FUNCTION_BLOCK "LModbusAscii_Master"   // FB4, SCL
TITLE = LModbusAscii_Master
{ S7_Optimized_Access := 'TRUE' }
AUTHOR : Siemens
FAMILY : LModbus
NAME : LModbusAscii_Master
VERSION : 1.1
// Modbus ASCII Master block
// the block implements the Modbus Ascii Master functionality
// ENO is not used, error handling done with error and status
   VAR_INPUT
      enable : Bool;   // True: Enables block functionality, rising edge initializes the port
      execute : Bool;   // Rising edge starts action once
      hardwareId : Hw_Any;   // Hardware Identifier for used communication module
      slaveAddress : USInt;   // Address of modbus ASCII Slave
      functionCode : USInt;   // Function code to send to the Slave
      startAddress : UInt;   // Startaddress in Modbus slave to read or write / if MB function 08, then startAddress is subfunctioncode / if MB function 43, then startAddress is object ID
      quantity : UInt;   // Quantity of Coils/Registers to read or write to /from slave device
      parameter : "LModbusAscii_typeAsciiConfiguration";   // Parameter dataset to configure modbus interface
      mask : Struct   // Logical Mask for Function Code 22 Mask Write Register
         andMask : Word;   // AND Mask of Function Code 22
         orMask : Word;   // OR Mask of Function Code 22
      END_STRUCT;
      readWrite : Struct   // Addresses and Quantities for Function Code 23 Read/Write Multiple registers
         startAddressRead : UInt := 1;   // Address to Holding Register for Read access
         quantityRead : USInt;   // Quantity of Holding Register for Read access
         startAddressWrite : UInt := 1;   // Address to Holding Register for Write access
         quantityWrite : USInt;   // Quantity of Holding Register for Write access
      END_STRUCT;
   END_VAR
   VAR_OUTPUT
      valid : Bool;   // TRUE: Valid set of output values available at the FB
      done : Bool;   // TRUE: Commanded functionality has been completed successfully
      busy : Bool;   // TRUE: FB is not finished and new output values can be expected
      error : Bool;   // TRUE: An error occurred during the execution of the FB
      status : Word := 16#7000;   // 16#0000 - 16#7FFF: Status of the FB, 16#8000 - 16#FFFF: Error identification
      diagnostics : "LModbusAscii_typeDiagnostics";   // Diagnostics information (status, subFunctionStatus, statenumber of Error)
   END_VAR
   VAR_IN_OUT
      data : Variant;   // Data for Modbus Read or Write of type Byte, Char, USInt, SInt, Bool, Word, UInt, Real, Int
   END_VAR
   VAR
      statExecuteOld : Bool;   // Old value of 'execute' input for edge detection
      statValid : Bool;   // Static value for output 'valid'
      statDone : Bool;   // Static value for output 'done'
      statBusy : Bool;   // Static value for output 'busy'
      statError : Bool;   // Static value for output 'error'
      statSerialLineStopBits : UInt;   // Serial line stop bits - defined by the parity
      statRetryCounter : USInt;   // Retry counter tag
      statFBState : DInt := 0;   // State in the state machine of the FB
      statDiagnostics : "LModbusAscii_typeDiagnostics";   // Static Diagnostic data and Information
      statEmptyDiagnostics : "LModbusAscii_typeDiagnostics";   // Empty diagnostics information (for initialization purposes only)
      statParameter : "LModbusAscii_typeAsciiConfiguration";
      instPortConfig : Port_Config;   // Instance Port configuration for Modbus ASCII Communication
      instTransmitterConfig : Send_Config;   // Instance Transmitter configuration for Modbus ASCII Communication
      instReceiverConfig : Receive_Config;   // Instance Receiver configuration for Modbus ASCII Communication
      statReceiverConditions : Receive_Conditions;   // Static Receive conditions for Modbus ASCII Communication
      instSendRequest : Send_P2P;   // Instance Send Data to Modbus slave
      instGetResponse : Receive_P2P;   // Instance Recive data from Modbus slave
      instResetRxBuffer : Receive_Reset;   // Instance Reset and clear receive buffer
      instWatchdog : IEC_TIMER;   // Instance Watchdog to check transmit to recive transition OR TurnAround delay time
      statTransmitterBuffer : Array[0..#BUFFER_UPPER_BOUND_BINARY] of Byte;   // Static Buffer for transmit data to slave device
      statReceiverBuffer : Array[0..#BUFFER_UPPER_BOUND_BINARY] of Byte;   // Static Buffer for receiving data from slave device
      statTransmitterAsciiBuffer : Array[0..#BUFFER_UPPER_BOUND_ASCII] of Byte;   // Static Buffer for the ASCII transfer string - send an receive direction
      statReceiverAsciiBuffer : Array[0..#BUFFER_UPPER_BOUND_ASCII] of Byte;   // Static Buffer for the ASCII transfer string - send an receive direction
      instAsciiDecode : "LModbusAscii_DecodeAsciiToByte";   // Instance to convert/decode the two ASCII nibble character array into byte array
      instAsciiEncode : "LModbusAscii_EncodeByteToAscii";   // Instance to convert/encode the byte array into a two ASCII nibble character array
      statReadWrite : Struct   // Addresses and Quantities for Function Code 23 Read/Write Multiple registers
         startAddressRead : UInt;
         quantityRead : USInt;
         startAddressWrite : UInt;
         quantityWrite : USInt;
      END_STRUCT;
      statHardwareId : UInt;   // Hardware Identifier for used communication module
      statErrorUserCleared : Bool;   // Error occurred that can only be solved by user; rising edge at enable input necessary
      statDisablingCompleted : Bool;   // TRUE: Disabling has been completed
      statErrorAutoCleared : Bool;   // Error occurred that can be acknowledged by FB
      statEnableOld : Bool;   // Old value of 'enable' input for edge detection
      statQuantityInBytes : USInt;   // Static internal value for quantity check in bytes
      statQuantityInBytesRead : USInt;   // Static internal value for quantity check in bytes for FC 23 Read requests
      statQuantityInBytesWrite : USInt;   // Static internal value for quantity check in bytes for FC 23 Write requests
      statFunctionCode : USInt;   // Function code to send to the Slave
      statSlaveAddress : USInt;   // Address of modbus ASCII Slave
      statQuantity : UInt;   // Static tag for quantity of requested data
      statStartAddress : UInt;   // Static tag for start address as word
      statAndMask : Word;   // AND Mask of Function Code 22
      statOrMask : Word;   // OR Mask of Function Code 22
      statLengthAfterEncoding : DInt;   // Temporary value for length of ASCII characters to transfer
      statLengthAfterDecoding : DInt;   // Temporary value for length of Byte Array received
   END_VAR
   VAR_TEMP
      tempExecute : Bool;   // Temporary value for input 'execute'
      tempStayInStatemachine : Bool;   // Temporary bool tag to stay in state machine and repeat execution if set to TRUE
      tempEnable : Bool;   // Temporary value for input 'enable'
      tempRetVal : Int;   // Temporary value for retVal of MOVE_BLK_VARIANT or DESERIALIZE
      tempSerializePos : DInt;   // Temporary value for serialize position
      tempDeserializePos : DInt;   // Temporary value for deserialize position
      tempReceiveBufferIndex : Int;   // Temporary value for receive buffer index
      tempLengthIndex : DInt;   // Temporary value for indexing buffer arrays
      tempEmptyData : Array[0..#BUFFER_UPPER_BOUND_BINARY] of Byte;   // Temporary value for reset data after disabling
      tempStartAddress : Word;   // Temporary value for Startaddress in Modbus slave to read or write / if MB function 08, then startAddress is subfunctioncode / if MB function 43, then startAddress is object ID
      tempQuantity : Word;   // Temporary value for Quantity of Coils/Registers to read or write to /from slave device
   END_VAR
   VAR CONSTANT
      FB_STATE_NO_PROCESSING_IDLE : DInt := 0;   // FB state: No processing
      FB_STATE_INIT_INTERFACE : DInt := 1;   // FB state: initialization of Port
      FB_STATE_INIT_TRANSMITTER : DInt := 2;   // FB state: initialization of Transmitter
      FB_STATE_INIT_RECEIVER : DInt := 3;   // FB state: initialization of Receiver
      FB_STATE_WAIT_FOR_EXECUTE : DInt := 4;   // FB state: wait until function should be executed
      FB_STATE_RESET_RECEIVER_BUFFER : DInt := 5;   // FB state: initialization of Receiver Buffer by clearing it
      FB_STATE_SETUP_TRANSMIT_PROTOCOL : DInt := 30;   // FB state: setup transmit protocol
      FB_STATE_TRANSMIT_DATA : DInt := 40;   // FB state: send message to slave
      FB_STATE_WAIT_FOR_RESPONSE : DInt := 41;   // FB state: wait for response from slave
      FB_STATE_WAIT_FOR_TURNAROUND_DELAY : DInt := 42;   // FB state: wait for turnaround delay after send broadcast
      FB_STATE_PROCESS_RECEIVED_DATA : DInt := 50;   // FB state: read / decode received data
      FB_STATE_DISABLING : DInt := 99;   // FB state: disabling / clear of the interface configuration
      STATUS_DONE : Word := 16#0000;   // Execution finished without errors
      STATUS_NO_CALL : Word := 16#7000;   // No job being currently processed
      STATUS_FIRST_CALL : Word := 16#7001;   // First call after enabling the block (rising edge 'enable')
      STATUS_SUBSEQUENT_CALL : Word := 16#7002;   // Subsequent call during active interface preparation without further details
      STATUS_READY : Word := 16#7003;   // Block is in ready state and waiting for a modbus job
      STATUS_EXECUTED_FIRST_CALL : Word := 16#7004;   // First call after incoming new job (rising edge 'execute')
      STATUS_EXECUTED_SUBSEQUENT_CALL : Word := 16#7005;   // Subsequent call during active job processing without further details
      NO_ERROR : Word := 16#0000;   // Blank error code / no error
      ERR_UNDEFINED_STATE : Word := 16#8600;   // Error due to an undefined state in state machine
      ERR_MODBUS_ADDRESS_OUT_OF_RANGE : Word := 16#8601;   // Error due to missconfiguration, Modbus address out of range 0 <= Address <= 247
      ERR_MODBUS_WRONG_PARITY_MODE : Word := 16#8602;   // Error due to missconfiguration, Modbus parity mode can be even(2), odd(3), no parity(1)
      ERR_MODBUS_WRONG_INTERFACE_MODE : Word := 16#8603;   // Error due to missconfiguration, Serial interface mode can be serial interface mode 0/FullDuplex (RS232), 4/Half duplex (RS485, two-wire mode)
      ERR_CONFIGURATION_PORT : Word := 16#8604;   // Error due to Port configuration, please check subfunction status in Diagnostic
      ERR_CONFIGURATION_TRANSMITTER : Word := 16#8605;   // Error due to Transmitter configuration, please check subfunction status in Diagnostic
      ERR_CONFIGURATION_RECEIVER : Word := 16#8606;   // Error due to Receiver configuration, please check subfunction status in Diagnostic
      ERR_CLEAR_RECEIVER_BUFFER : Word := 16#8607;   // Error due to clear Receiver buffer, please check subfunction status in Diagnostic
      ERR_MOVE_BLK_VAR_TO_DATA : Word := 16#8608;   // Error due to moving received data to INOUT data
      ERR_DESERIALIZE_TO_DATA : Word := 16#8609;   // Error due to deserializing received data to INOUT data
      ERR_REQUEST_NOT_SUPPORTED_FUNCTION_CODE : Word := 16#8610;   // Error due to given Modbus Function Code, not supported function, see subFctStatus in diagnostic
      ERR_REQUEST_INVALID_FC08_REQUEST_DATA : Word := 16#8681;   // Error due to given request data - for function code 8 / sub function code 1 data field needs to be 16#0000 (leave log) or 16#FF00 (clear log)
      ERR_RESPONSE_NOT_SUPPORTED_FUNCTION_CODE : Word := 16#8620;   // Error due to received Modbus Function Code, not supported function, see subFctStatus in diagnostic
      ERR_INTERFACE_NOT_CONFIGURED : Word := 16#8611;   // Error due to interface, that was not configured yet
      ERR_SERIALIZE_MULTIPLE_WRITE : Word := 16#8612;   // Error due to serializing data to transmitter buffer at multiple write request
      ERR_SERIALIZE_SINGLE_WRITE : Word := 16#8622;   // Error due to serializing data to transmitter buffer at single write request
      ERR_MOVE_BLK_VAR_MULTIPLE_WRITE : Word := 16#8613;   // Error due to moving data to transmitter buffer
      ERR_INVALID_QUANTITY : Word := 16#8615;   // Error due to invalid quantity for read (125) or write (121) request
      ERR_MOVE_BLK_VAR_RECEIVE_DATA : Word := 16#8633;   // Error due to moving receive buffer to data
      ERR_MOVE_BLK_VAR_SINGLE_WRITE : Word := 16#8623;   // Error due to moving data to transmitter buffer
      ERR_DATA_TYPE_NOT_SUPPORTED : Word := 16#8614;   // Error due to moving data to INOUT data. Has to be Array of Byte or Word.
      ERR_TRANSMISSION_FAILURE : Word := 16#8201;   // Error during data transmisson to slave, please check subfunction status in Diagnostic
      ERR_RESPONSE_TIMEOUT_EXPIRATION : Word := 16#8202;   // Error due to timeout while wait for response from slave, "response time-out expiration"
      ERR_RECEIVER_FAILURE : Word := 16#8203;   // Error due to receiver data from slave, please check subfunction status in Diagnostic
      ERR_RESPONSE_EXCEPTION_FROM_SLAVE : Word := 16#8204;   // Error due to an received exception from slave - excpetion code is stored in diagnostics subFunctionStatus
      ERR_RESPONSE_WRONG_LRC : Word := 16#8205;   // Error due to LRC Check on response data
      ERR_RESPONSE_WRONG_QUANTITY : Word := 16#8206;   // Error due to wrong quantity received
      ERR_RESPONSE_SINGLE_WRITE : Word := 16#8207;   // Error due to response of single write functions
      ERR_RESPONSE_MULTI_WRITE : Word := 16#8217;   // Error due to response of multiple write functions
      ERR_RESPONSE_NOT_EXPECTED_FC : Word := 16#8208;   // Error because response contains not expected function code
      ERR_RESPONSE_NOT_EXPECTED_SUB_FC : Word := 16#8218;   // Error because response contains not expected subfunction code
      ERR_RESPONSE_WRONG_SLAVE : Word := 16#8209;   // Error due to wrong slave answered to request
      ERR_NOT_SUPPORTED_SUB_FC : Word := 16#8210;   // Error due to not supported function code for diagnostic function 08
      ERR_DIAG_SUB_0 : Word := 16#8250;   // Error in response for diagnostic subfunction 0 (Return query value) - wrong echo value
      ERR_DIAG_SUB_1 : Word := 16#8251;   // Error in response for diagnostic subfunction 1 (Restart Com) - wrong echo value
      FREEPORT_PROTOCOL : UInt := 0;   // Freeport protocol is used for Modbus ASCII
      FB_DISABLE_TIME : Time := T#500Ms;   // Time that any active instances may need until the device is hard deactivated.
      BUFFER_UPPER_BOUND_ASCII : DInt := 608;   // Upper Bound of Buffer ASCII Char mode
      BUFFER_UPPER_BOUND_BINARY : DInt := 300;   // Upper Bound of Buffer in Byte to store the binary data
      DATA_INDEX_0 : Int := 0;   // Data index set to 0
      INITIALIZE_WORD_0 : Word := 16#0000;   // Initialize Word (16#00)
      B1_OFFSET : USInt := 1;   // Offset to select high byte in a word
      FC05_SET_COMMAND_IDENT : Word := 16#FF00;   // Modbus ASCII - identifier for setting coil to true
      MODBUS_INTERFACE_MODE_RS232 : USInt := 0;   // Modbus interface modus is RS232 Full Duplex
      MODBUS_INTERFACE_MODE_RS485 : USInt := 4;   // Modbus interface modus is RS485 Half Duplex
      MODBUS_ADDRESS_MAX : USInt := 247;   // Modbus ASCII maximum address range is 247
      MODBUS_ADDRESS_BROADCAST : USInt := 0;   // Modbus ASCII broadcast address is 0
      MODBUS_ASCII_SEVEN_DATABITS : UInt := 2;   // Modbus ASCII Databits defined --> 7
      MODBUS_ASCII_PARITY_EVEN : UInt := 2;   // Modbus ASCII EVEN Parity setting for port configuration
      MODBUS_ASCII_PARITY_ODD : UInt := 3;   // Modbus ASCII ODD Parity setting for port configuration
      MODBUS_ASCII_NO_PARITY : UInt := 1;   // Modbus ASCII NO Parity setting for port configuration
      MODBUS_ASCII_STOPBITS_NO_PARITY : UInt := 2;   // Modbus ASCII Stopbits = 2 if no parity mode is choosen
      MODBUS_ASCII_STOPBITS_WITH_PARITY : UInt := 1;   // Modbus ASCII Stopbits = 1 if even or odd parity mode is choosen
      MODBUS_TURNAROUND_DELAY : Time := T#200MS;   // Modbus turnaround delay time after a broadcast request was send
      MODBUS_SLAVE_ADDRESS_INDEX : USInt := 0;   // Modbus Master / Slave request / response - index for slave address
      MODBUS_FUNCTION_CODE_INDEX : USInt := 1;   // Modbus Master / Slave request / response - index for function code AND Exception notice (MSB) in response buffer
      MODBUS_RESPONSE_BYTE_COUNT_INDEX : USInt := 2;   // Modbus Master - Index to length entry in response field
      MODBUS_RESPONSE_ADDRESS_INDEX : USInt := 2;   // Modbus Master - Index to start address in response field
      MODBUS_RESPONSE_QUANTITY_INDEX : USInt := 4;   // Modbus Master - Index to quantity in response field
      MODBUS_EXCEPTION_CODE_INDEX : USInt := 1;   // Modbus Slave response - index for exception code in response buffer
      MODBUS_DEFAULT_REQUEST_LENGTH : USInt := 2;   // Modbus Master request - shortest possible request length
      MODBUS_DEFAULT_RESP_INDEX : USInt := 2;   // Modbus Master response - default response index
      MODBUS_STARTADDRESS_INDEX : USInt := 2;   // Modbus Master request - index for start address
      MODBUS_STARTADDRESS_FC23_WRITE_INDEX : USInt := 6;   // Modbus Master request - index for start address of write job for FC 23 request
      MODBUS_AND_MASK_INDEX : USInt := 4;   // Modbus Master request - index for AND Mask for fc 22
      MODBUS_OR_MASK_INDEX : USInt := 6;   // Modbus Master request - index for OR Mask for fc 22
      MODBUS_QUANTITY_INDEX : USInt := 4;   // Modbus Master request - index for quantity
      MODBUS_QUANTITY_FC23_WRITE_INDEX : USInt := 8;   // Modbus Master request - index for quantity of write job for FC 23 request
      MODBUS_BYTE_COUNT_INDEX : USInt := 6;   // Modbus Master request - index byte count
      MODBUS_BYTE_COUNT_FC23_INDEX : USInt := 10;   // Modbus Master request - index byte count of write job for FC 23 request
      MODBUS_DATA_INDEX : USInt := 7;   // Modbus Master request - index to first data entry
      MODBUS_FC23_DATA_INDEX : USInt := 11;   // Modbus Master request - index to first data entry of write job for FC 23 request
      MODBUS_USER_DATA_READ_INDEX : USInt := 3;   // Modbus Slave response - index for position of user data
      MODBUS_DIAG_SUB_FC_INDEX : USInt := 2;   // Modbus Master / Slave request / Response - index for subfunction code at Diagnostic function and Device ident
      MODBUS_DIAG_DATA_INDEX : USInt := 4;   // Modbus Master / Slave request / Response - index for subfunction code at Diagnostic function and Device ident
      MODBUS_REQUEST_LENGTH : UInt := 6;   // Modbus Master request length
      MODBUS_REQUEST_MULTIPLE_WRITE_LENGTH : UInt := 7;   // Modbus Master request length for multiple write functions
      MODBUS_REQUEST_MASK_WRITE_LENGTH : UInt := 8;   // Modbus Master request length for mask write function
      MODBUS_REQUEST_READ_WRITE_LENGTH : UInt := 11;   // Modbus Master request length for FC 23 read/write request
      MODBUS_STARTADDRESS_CORRECTION : USInt := 1;   // Correction of MODBUS startaddress by subtraction of 1
      MODBUS_MAX_REGISTER_READ : USInt := 125;   // Modbus maximum quantity for register read requests
      MODBUS_MAX_REGISTER_WRITE : USInt := 123;   // Modbus maximum quantity for register write requests
      MODBUS_FC23_MAX_REGISTER_WRITE : USInt := 121;   // Modbus maximum quantity for FC 23 register write requests
      MODBUS_FC43_MEI_TYE : Byte := 16#0E;   // Modbus MEI Type for Device Identification
      MODBUS_FC43_DEVICE_ID_CODE_INDEX : USInt := 3;   // Modbus Device ID code index in request
      MODBUS_FC43_OBJECT_ID_CODE_INDEX : USInt := 4;   // Modbus Object ID code index in request
      MODBUS_FC43_REQUEST_LENGTH : USInt := 5;   // Modbus Master request length for FC 43 request
      MB_FC_01_READ_COILS : USInt := 1;   // Modbus function code 01 - read coils
      MB_FC_02_READ_DISCRETE_INPUTS : USInt := 2;   // Modbus function code 02 - read discrete inputs
      MB_FC_03_READ_HOLDING_REGISTERS : USInt := 3;   // Modbus function code 03 - read holding registers
      MB_FC_04_READ_INPUT_REGISTERS : USInt := 4;   // Modbus function code 04 - read input registers
      MB_FC_05_WRITE_COIL : USInt := 5;   // Modbus function code 05 - write single coil
      MB_FC_06_WRITE_REGISTER : USInt := 6;   // Modbus function code 06 - write single register
      MB_FC_07_READ_EXCEPTION_STATUS : USInt := 7;   // Modbus function code 07 - read exception status
      MB_FC_08_DIAGNOSTIC : USInt := 8;   // Modbus function code 08 - diagnostic
      MB_FC_11_GET_COM_EVENT_COUNTER : USInt := 11;   // Modbus function code 11 - diagnostic
      MB_FC_12_GET_COM_EVENT_LOG : USInt := 12;   // Modbus function code 12 - get comm event log
      MB_FC_15_WRITE_COILS : USInt := 15;   // Modbus function code 15 - write multiple coils
      MB_FC_16_WRITE_REGISTERS : USInt := 16;   // Modbus function code 16 - write multiple registers
      MB_FC_22_MASK_WRITE_REGISTER : USInt := 22;   // Modbus function code 22 - mask Write Register
      MB_FC_23_READ_WRITE_MULTIPLE_REGISTERS : USInt := 23;   // Modbus function code 23 - read/write Multiple registers
      MB_FC_43_READ_DEVICE_IDENT : USInt := 43;   // Modbus function code 43 - read device idendification data
      DIAG_SUB_FC_0_RETURN_QUERY_DATA : USInt := 16#00;   // Diag: Return query dara
      DIAG_SUB_FC_1_RESTART_COM : USInt := 16#01;   // Diag: Restart communication option
      DIAG_SUB_FC_2_RETURN_DIAG_REGISTER : USInt := 16#02;   // Diag: Return diagnostic register
      DIAG_SUB_FC_4_FORCE_LISTEN_ONLY : USInt := 16#04;   // Diag: Force listen only
      DIAG_SUB_FC_10_CLEAR_DIAG_REGISTER : USInt := 16#0A;   // Diag: Clear counter and diagnostic register
      DIAG_SUB_FC_11_COUNTER_TOTAL_MESSAGE : USInt := 16#0B;   // Diag: Return bus message count
      DIAG_SUB_FC_12_COUNTER_CRC_ERR : USInt := 16#0C;   // Diag: Return bus commuunication error count
      DIAG_SUB_FC_13_COUNTER_EXCEPTION_ERR : USInt := 16#0D;   // Diag: Return bus exception error count
      DIAG_SUB_FC_14_COUNTER_TOTAL_MESSAGES : USInt := 16#0E;   // Diag: Return server message count
      DIAG_SUB_FC_15_COUNTER_NO_RESPONSE : USInt := 16#0F;   // Diag: Return Server no respomse count
      DIAG_SUB_FC_16_COUNTER_NAK : USInt := 16#10;   // Diag: Return Server negative acknowledge count
      DIAG_SUB_FC_17_COUNTER_SERVER_BUSY : USInt := 16#11;   // Diag: Return Server busy count
      DIAG_SUB_FC_18_BUS_CHAR_OVERRUN : USInt := 16#12;   // Diag: Return Bus Character Overrun Count
      DIAG_SUB_FC_20_CLEAR_OVERRUN : USInt := 16#14;   // Diag: Clear Overrun Counter and Flag
   END_VAR
   // statDiagnostics.status := 16#7000;
BEGIN
   REGION BLOCK INFO HEADER
     //===============================================================================
     // SIEMENS / (c)copyright 2026
     //-------------------------------------------------------------------------------
     // Title:            LModbusAscii_Master
     // Comment/Function: Modbus ASCII Master
     //                   The block implements the Modbus ASCII Master functionality.
     //                   ENO is not used, error handling done with error and status.
     // Library/Family:   LModbus
     // Author:           Siemens
     // Tested with:      S7-1200/1500
     // Engineering:      TIA Portal >= V19
     // Restrictions:     (none)
     // Requirements:     CM (RS485)
     //-------------------------------------------------------------------------------
     // Change log table:
     // Version  | Date       | Expert in charge       | Changes applied
     //----------|------------|------------------------|------------------------------
     // 00.01.00 | 2019-08-05 | Siemens                | first released version
     // 01.00.00 | 2023-03-20 | Siemens                | Styleguide adaptions and bugfix for data output
     // 01.01.00 | 2026-05-29 | Siemens                | New Functions and BugFix
     //===============================================================================
   END_REGION

   REGION ENABLING/DISABLING
     #tempEnable := #enable; // work with temporary value
     #tempExecute := #execute; // work with temporary value

     IF (#tempEnable = TRUE) AND (#statDiagnostics.status = #STATUS_NO_CALL) THEN // Enable FB
       REGION Enable
         // first call; initialize FB
         REGION Initialize standard interface
           #statBusy := TRUE;
           #statError := FALSE;
           #statErrorUserCleared := FALSE;
           #statErrorAutoCleared := FALSE;
           #statDiagnostics.status := #STATUS_FIRST_CALL;
           #statDiagnostics.subFunctionStatus := #NO_ERROR;
           #statDiagnostics.stateNumber := 0;
           #diagnostics := #statEmptyDiagnostics;
           #statDisablingCompleted := FALSE;
         END_REGION Initialize standard interface

         REGION Verify Input parameters
           #statParameter := #parameter;
           // verify interface mode is RS232 or RS485
           IF #statParameter.modeInterfacePTP <> #MODBUS_INTERFACE_MODE_RS232
             AND #statParameter.modeInterfacePTP <> #MODBUS_INTERFACE_MODE_RS485
           THEN
             #statErrorUserCleared := TRUE;
             #statDiagnostics.status := #ERR_MODBUS_WRONG_INTERFACE_MODE;

             // check parity mode even odd or non parity
           ELSIF #statParameter.parity <> #MODBUS_ASCII_NO_PARITY
             AND #statParameter.parity <> #MODBUS_ASCII_PARITY_EVEN
             AND #statParameter.parity <> #MODBUS_ASCII_PARITY_ODD
           THEN
             #statErrorUserCleared := TRUE;
             #statDiagnostics.status := #ERR_MODBUS_WRONG_PARITY_MODE;
           END_IF;

           #statHardwareId := #hardwareId;
         END_REGION

         REGION Init static tags
           // adjust stop bits for serial interface configuration
           IF #statParameter.parity = #MODBUS_ASCII_NO_PARITY THEN
             // if no Parity is choosen, two stop bits are needed
             #statSerialLineStopBits := #MODBUS_ASCII_STOPBITS_NO_PARITY;
           ELSE
             // if even or odd Parity is choosen, just one stop bit is needed
             #statSerialLineStopBits := #MODBUS_ASCII_STOPBITS_WITH_PARITY;
           END_IF;
         END_REGION Init static tags

         REGION Init instances by call subsidiary FBs with false
           #instPortConfig(REQ := FALSE);
           #instTransmitterConfig(REQ := FALSE);
           #instReceiverConfig(REQ := FALSE,
                               Receive_Conditions := #statReceiverConditions);
           #instSendRequest(REQ := FALSE,
                            BUFFER:=#statTransmitterAsciiBuffer);
         END_REGION Init instances by call subsidiary FBs with false

         // state machine - start functionality
         #statFBState := #FB_STATE_INIT_INTERFACE;
       END_REGION Enable

     ELSIF (#tempEnable = FALSE) AND (#statEnableOld = TRUE) THEN // disable FB 
       REGION Disable
         #statFBState := #FB_STATE_DISABLING;
         #instWatchdog.TON(IN := FALSE, PT := #FB_DISABLE_TIME);
       END_REGION Disable

     ELSIF (#statDiagnostics.status = #STATUS_FIRST_CALL) THEN // set status identifier of subsequent call
       REGION Subsequent
         #statDiagnostics.status := #STATUS_SUBSEQUENT_CALL;
       END_REGION Subsequent

     ELSIF NOT #tempEnable
       AND #statDiagnostics.status = #STATUS_NO_CALL
       AND (#tempExecute = TRUE)
       AND (#statExecuteOld = FALSE) // check if FB is triggered
     THEN
       REGION Faulty Call - execute with disabled function block
         #statErrorUserCleared := TRUE;
         #statDiagnostics.status := #ERR_INTERFACE_NOT_CONFIGURED;
         #statDiagnostics.subFunctionStatus := #NO_ERROR;
       END_REGION Faulty Call - execute with disabled function block

     END_IF;

     // edge detection 'enable' input
     #statEnableOld := #tempEnable;
   END_REGION ENABLING/DISABLING

   IF (#statDiagnostics.status = #STATUS_NO_CALL) THEN // nothing to do -> End here to reduce "system load"
     RETURN;
   END_IF;

   REGION STATE_MACHINE
     REPEAT
       // set repeat condition to FALSE to leave state machine loop
       #tempStayInStatemachine := FALSE;
       CASE #statFBState OF // state machine of FB
         #FB_STATE_NO_PROCESSING_IDLE: // no processing active (Note: this state must always be present and left empty)
           REGION No Processing
             ;
           END_REGION No Processing

         #FB_STATE_INIT_INTERFACE:
           REGION Init Interface
             // call port configuration to set parameters for communication
             #instPortConfig(REQ := TRUE,
                             "PORT" := #statHardwareId,
                             PROTOCOL := #FREEPORT_PROTOCOL,
                             BAUD := #statParameter.baud,
                             PARITY := #statParameter.parity,
                             DATABITS := #MODBUS_ASCII_SEVEN_DATABITS,
                             STOPBITS := #statSerialLineStopBits,
                             MODE := #statParameter.modeInterfacePTP);

             // port configuration finished successfully
             IF (#instPortConfig.DONE = TRUE) THEN
               #instPortConfig(REQ := FALSE);  // reset port config REQ input after call
               #statFBState := #FB_STATE_INIT_TRANSMITTER;   // set next state

               // error occurred during Port Configuration
             ELSIF (#instPortConfig.ERROR = TRUE) THEN
               // write diagnostic Information
               #statErrorUserCleared := TRUE;
               #statDiagnostics.status := #ERR_CONFIGURATION_PORT; // set correct status that identifies error clearly
               #statDiagnostics.subFunctionStatus := #instPortConfig.STATUS; // status of Port Configuration
               #statDiagnostics.stateNumber := #statFBState; // set error state number for diagnostic

               #instPortConfig(REQ := FALSE); // reset port config REQ input after call
             END_IF;
           END_REGION Init Interface

         #FB_STATE_INIT_TRANSMITTER:
           REGION Init Transmitter
             // call transmitter configuration to set paramters for communication (SEND_CFG)
             #instTransmitterConfig(REQ := TRUE,
                                    "PORT" := #statHardwareId);

             // port configuration finished successfully
             IF (#instTransmitterConfig.DONE = TRUE) THEN
               #instTransmitterConfig(REQ := FALSE);   // reset receiver config REQ input after call
               #statFBState := #FB_STATE_INIT_RECEIVER;  // set next state

               // error occurred during Port Configuration
             ELSIF (#instTransmitterConfig.ERROR = TRUE) THEN
               // write diagnostic Information
               #statErrorUserCleared := TRUE;
               #statDiagnostics.status := #ERR_CONFIGURATION_TRANSMITTER; // set correct status that identifies error clearly
               #statDiagnostics.subFunctionStatus := #instTransmitterConfig.STATUS; // status of Port Configuration
               #statDiagnostics.stateNumber := #statFBState; // set error state number for diagnostic

               #instTransmitterConfig(REQ := FALSE); // reset receiver config REQ input after call
             END_IF;
           END_REGION Init Transmitter

         #FB_STATE_INIT_RECEIVER:
           REGION Init Receiver
             // call receiver configuration to set paramters for communication (RCV_CFG)
             #instReceiverConfig(REQ := TRUE,
                                 "PORT" := #statHardwareId,
                                 Receive_Conditions := #statReceiverConditions);

             // port configuration finished successfully
             IF (#instReceiverConfig.DONE = TRUE) THEN
               #instReceiverConfig(REQ := FALSE,
                                   Receive_Conditions := #statReceiverConditions); // reset receiver config REQ input after call

               #statValid := TRUE;
               #statBusy := FALSE;
               #statDiagnostics.status := #STATUS_READY;
               #statFBState := #FB_STATE_WAIT_FOR_EXECUTE; // set next state

               // error occurred during Port Configuration
             ELSIF (#instReceiverConfig.ERROR = TRUE) THEN
               // write diagnostic Information
               #statErrorUserCleared := TRUE;
               #statDiagnostics.status := #ERR_CONFIGURATION_RECEIVER; // set correct status that identifies error clearly
               #statDiagnostics.subFunctionStatus := #instReceiverConfig.STATUS; // status of Port Configuration
               #statDiagnostics.stateNumber := #statFBState; // set error state number for diagnostic

               #instReceiverConfig(REQ := FALSE,
                                   Receive_Conditions := #statReceiverConditions); // reset receiver config REQ input after call
             END_IF;
           END_REGION Init Receiver

         #FB_STATE_WAIT_FOR_EXECUTE:
           REGION Wait for execute
             REGION Execute
               IF (#tempExecute = TRUE) AND (#statExecuteOld = FALSE) // check if FB is triggered
               THEN
                 REGION Verify input paramters
                   #statFunctionCode := #functionCode;
                   #statSlaveAddress := #slaveAddress;

                   // check, if requested function code is supported by the function block
                   IF #statFunctionCode <> #MB_FC_01_READ_COILS
                     AND #statFunctionCode <> #MB_FC_02_READ_DISCRETE_INPUTS
                     AND #statFunctionCode <> #MB_FC_03_READ_HOLDING_REGISTERS
                     AND #statFunctionCode <> #MB_FC_04_READ_INPUT_REGISTERS
                     AND #statFunctionCode <> #MB_FC_05_WRITE_COIL
                     AND #statFunctionCode <> #MB_FC_06_WRITE_REGISTER
                     AND #statFunctionCode <> #MB_FC_07_READ_EXCEPTION_STATUS
                     AND #statFunctionCode <> #MB_FC_08_DIAGNOSTIC
                     AND #statFunctionCode <> #MB_FC_11_GET_COM_EVENT_COUNTER
                     AND #statFunctionCode <> #MB_FC_12_GET_COM_EVENT_LOG
                     AND #statFunctionCode <> #MB_FC_15_WRITE_COILS
                     AND #statFunctionCode <> #MB_FC_16_WRITE_REGISTERS
                     AND #statFunctionCode <> #MB_FC_22_MASK_WRITE_REGISTER
                     AND #statFunctionCode <> #MB_FC_23_READ_WRITE_MULTIPLE_REGISTERS
                     AND #statFunctionCode <> #MB_FC_43_READ_DEVICE_IDENT
                   THEN
                     REGION invalid function code
                       // FB stays in wait for execute state and can be triggerde again with supported function code
                       #statErrorAutoCleared := TRUE;
                       #statDiagnostics.status := #ERR_REQUEST_NOT_SUPPORTED_FUNCTION_CODE;
                       #statDiagnostics.subFunctionStatus := USINT_TO_WORD(#statFunctionCode); // Given function code
                       #statDiagnostics.stateNumber := #statFBState; // Set error state number for diagnostic
                       EXIT; //end of block
                     END_REGION invalid function code

                   ELSIF #statSlaveAddress > #MODBUS_ADDRESS_MAX THEN
                     REGION invalid slave address
                       // verify Modbus address exceeds maximum address range
                       #statErrorAutoCleared := TRUE;
                       #statDiagnostics.subFunctionStatus := USINT_TO_WORD(#statSlaveAddress);
                       #statDiagnostics.status := #ERR_MODBUS_ADDRESS_OUT_OF_RANGE;
                       #statDiagnostics.stateNumber := #statFBState;
                       EXIT;
                     END_REGION invalid slave address

                   ELSE
                     REGION initialize function code
                       // set internal retry counter
                       // copy number of retries for retry transmition counter
                       #statRetryCounter := #statParameter.numberOfRetries;

                       // initialize statQuantity and statStartAddress
                       #statQuantity := #quantity;
                       #statStartAddress := #startAddress;

                       // check requested quantity. Later this value will be compared with the received data
                       IF #statFunctionCode = #MB_FC_01_READ_COILS
                         OR #statFunctionCode = #MB_FC_02_READ_DISCRETE_INPUTS
                         OR #statFunctionCode = #MB_FC_15_WRITE_COILS
                       THEN
                         //parameter quantity means count of bits. Eight bits are one bytes long
                         #statQuantityInBytes := UINT_TO_USINT(#statQuantity / 8);
                         IF #statQuantity MOD 8 <> 0 THEN
                           #statQuantityInBytes += 1;
                         END_IF;

                       ELSIF #statFunctionCode = #MB_FC_03_READ_HOLDING_REGISTERS
                         OR #statFunctionCode = #MB_FC_04_READ_INPUT_REGISTERS
                         OR #statFunctionCode = #MB_FC_16_WRITE_REGISTERS
                       THEN
                         // parameter quantity means count of registers. One register is two bytes long
                         #statQuantityInBytes := UINT_TO_USINT(#statQuantity) * 2;

                       ELSIF (#statFunctionCode = #MB_FC_08_DIAGNOSTIC AND #statQuantity <> #DIAG_SUB_FC_4_FORCE_LISTEN_ONLY)
                         OR #statFunctionCode = #MB_FC_05_WRITE_COIL
                         OR #statFunctionCode = #MB_FC_06_WRITE_REGISTER
                         OR #statFunctionCode = #MB_FC_07_READ_EXCEPTION_STATUS
                       THEN
                         // two bytes fixed for reply request (ping behaviour) and for single register and coil write 
                         #statQuantityInBytes := 2;

                       ELSIF #statFunctionCode = #MB_FC_22_MASK_WRITE_REGISTER THEN
                         #statQuantityInBytes := 0;
                         #statAndMask := #mask.andMask;
                         #statOrMask := #mask.orMask;

                       ELSIF #statFunctionCode = #MB_FC_23_READ_WRITE_MULTIPLE_REGISTERS THEN
                         #statReadWrite.startAddressRead := #readWrite.startAddressRead;
                         #statReadWrite.quantityRead := #readWrite.quantityRead;
                         #statReadWrite.startAddressWrite := #readWrite.startAddressWrite;
                         #statReadWrite.quantityWrite := #readWrite.quantityWrite;
                         #statQuantityInBytesRead := #statReadWrite.quantityRead * 2;
                         #statQuantityInBytesWrite := #statReadWrite.quantityWrite * 2;

                       ELSIF #statFunctionCode = #MB_FC_11_GET_COM_EVENT_COUNTER THEN
                         #statQuantityInBytes := 4;

                       ELSIF #statFunctionCode = #MB_FC_43_READ_DEVICE_IDENT THEN
                         #statQuantityInBytes := 250;
                       END_IF;
                     END_REGION initialize function code

                   END_IF;

                 END_REGION Verify input paramters

                 REGION Init instances by call subsidiary FBs with FALSE
                   #instResetRxBuffer(REQ := FALSE,
                                      "PORT" := #statHardwareId);
                   #instWatchdog.TON(IN := FALSE,
                                     PT := #statParameter.transmissionWatchdog);
                 END_REGION Init instances by call subsidiary FBs with FALSE

                 // state machine - start processing
                 #statBusy := TRUE;
                 #statFBState := #FB_STATE_RESET_RECEIVER_BUFFER;
                 #statDiagnostics.status := #STATUS_EXECUTED_FIRST_CALL;

               ELSIF NOT #tempExecute AND #statDone THEN
                 #statDiagnostics.status := #STATUS_READY;
                 #statDone := FALSE;
                 #statError := FALSE;
               END_IF;

               // edge detection 'execute' input
               #statExecuteOld := #tempExecute;
             END_REGION Execute
           END_REGION

         #FB_STATE_RESET_RECEIVER_BUFFER:
           REGION Reset Receiver Buffer
             IF #statDiagnostics.status = #STATUS_EXECUTED_FIRST_CALL THEN
               #statDiagnostics.status := #STATUS_EXECUTED_SUBSEQUENT_CALL;
             END_IF;

             // call receiver reset buffer to clear it
             #instResetRxBuffer(REQ := TRUE,
                                "PORT" := #statHardwareId);

             // port configuration finished successfully
             IF (#instResetRxBuffer.DONE = TRUE) THEN
               #instResetRxBuffer(REQ := FALSE);   // reset receiver config REQ input after call
               #statFBState := #FB_STATE_SETUP_TRANSMIT_PROTOCOL;  // set next state

               // error occurred during Port Configuration
             ELSIF (#instResetRxBuffer.ERROR = TRUE) THEN
               // write diagnostic Information
               #statErrorAutoCleared := TRUE;
               #statDiagnostics.status := #ERR_CLEAR_RECEIVER_BUFFER; // set correct status that identifies error clearly
               #statDiagnostics.subFunctionStatus := #instResetRxBuffer.STATUS; // status of Port Configuration
               #statDiagnostics.stateNumber := #statFBState; // set error state number for diagnostic

               #instResetRxBuffer(REQ := FALSE);   // reset receiver config REQ input after call
             END_IF;
           END_REGION Init Receiver Buffer

         #FB_STATE_SETUP_TRANSMIT_PROTOCOL:
           REGION Setup Transmit Protocol
             // set up communication Buffer
             // first part: is the address
             #statTransmitterBuffer[#MODBUS_SLAVE_ADDRESS_INDEX] := USINT_TO_BYTE(#statSlaveAddress);
             // second part: is the function code
             #statTransmitterBuffer[#MODBUS_FUNCTION_CODE_INDEX] := USINT_TO_BYTE(#statFunctionCode);
             // third part: set start address for request

             IF #statFunctionCode <> #MB_FC_08_DIAGNOSTIC AND #statFunctionCode <> #MB_FC_43_READ_DEVICE_IDENT THEN
               #statStartAddress := #statStartAddress - #MODBUS_STARTADDRESS_CORRECTION;
             END_IF;

             // third part: tx / transmit data protocol setup
             // depending on the function code
             REGION Setup function code specific part
               CASE #statFunctionCode OF

                 #MB_FC_01_READ_COILS,
                 #MB_FC_02_READ_DISCRETE_INPUTS:
                   REGION 01 / 02 Read Coils/Discrete Inputs
                     // write start address to array
                     #tempStartAddress := UINT_TO_WORD(#statStartAddress);
                     #statTransmitterBuffer[#MODBUS_STARTADDRESS_INDEX] := #tempStartAddress.%B1;
                     #statTransmitterBuffer[#MODBUS_STARTADDRESS_INDEX + #B1_OFFSET] := #tempStartAddress.%B0;

                     // write quantity to array
                     #tempQuantity := UINT_TO_WORD(#statQuantity);
                     #statTransmitterBuffer[#MODBUS_QUANTITY_INDEX] := #tempQuantity.%B1;
                     #statTransmitterBuffer[#MODBUS_QUANTITY_INDEX + #B1_OFFSET] := #tempQuantity.%B0;

                     #tempLengthIndex := #MODBUS_REQUEST_LENGTH;
                   END_REGION

                 #MB_FC_03_READ_HOLDING_REGISTERS,
                 #MB_FC_04_READ_INPUT_REGISTERS:
                   REGION 03 / 04 Read Holding/Input Registers
                     // write start address to array
                     #tempStartAddress := UINT_TO_WORD(#statStartAddress);
                     #statTransmitterBuffer[#MODBUS_STARTADDRESS_INDEX] := #tempStartAddress.%B1;
                     #statTransmitterBuffer[#MODBUS_STARTADDRESS_INDEX + #B1_OFFSET] := #tempStartAddress.%B0;

                     // write quantity to array
                     #tempQuantity := UINT_TO_WORD(#statQuantity);
                     #statTransmitterBuffer[#MODBUS_QUANTITY_INDEX] := #tempQuantity.%B1;
                     #statTransmitterBuffer[#MODBUS_QUANTITY_INDEX + #B1_OFFSET] := #tempQuantity.%B0;

                     // set request length for ASCII encoding
                     #tempLengthIndex := #MODBUS_REQUEST_LENGTH;
                   END_REGION

                 #MB_FC_05_WRITE_COIL,
                 #MB_FC_06_WRITE_REGISTER:
                   REGION 05 / 06 Write coil/Register
                     // write start address to array
                     #tempStartAddress := UINT_TO_WORD(#statStartAddress);
                     #statTransmitterBuffer[#MODBUS_STARTADDRESS_INDEX] := #tempStartAddress.%B1;
                     #statTransmitterBuffer[#MODBUS_STARTADDRESS_INDEX + #B1_OFFSET] := #tempStartAddress.%B0;

                     IF IS_ARRAY(#data) AND
                       (TypeOfElements(#data) = Byte OR TypeOfElements(#data) = Char)
                     THEN
                       // for an array at INOUT data MOVE_BLK_VARIANT is used to copy data from static receive buffer to the INOUT
                       #tempRetVal := MOVE_BLK_VARIANT(SRC := #data,
                                                       COUNT := #statQuantityInBytes,
                                                       SRC_INDEX := #DATA_INDEX_0,
                                                       DEST_INDEX := #MODBUS_QUANTITY_INDEX,
                                                       DEST => #statTransmitterBuffer);
                       // if MOVE_BLK_VARIANT was executed with error, jump to AutoCleard error and give feedback to the user
                       IF #tempRetVal <> 0 THEN
                         #statErrorAutoCleared := TRUE;
                         #statDiagnostics.status := #ERR_MOVE_BLK_VAR_SINGLE_WRITE;
                         #statDiagnostics.subFunctionStatus := INT_TO_WORD(#tempRetVal);
                         #statDiagnostics.stateNumber := #statFBState;
                       END_IF;

                     ELSE
                       // for a structure or other data type at INOUT data serialized is used to copy data from static receive buffer to the INOUT
                       #tempSerializePos := #MODBUS_QUANTITY_INDEX;
                       #tempRetVal := Serialize(SRC_VARIABLE := #data,
                                                DEST_ARRAY => #statTransmitterBuffer,
                                                POS := #tempSerializePos);
                       // if serialize function was executed with error, jump to AutoCleared error and give feedback to the user
                       IF #tempRetVal <> 0 THEN
                         #statErrorAutoCleared := TRUE;
                         #statDiagnostics.status := #ERR_SERIALIZE_SINGLE_WRITE;
                         #statDiagnostics.subFunctionStatus := INT_TO_WORD(#tempRetVal);
                         #statDiagnostics.stateNumber := #statFBState;
                       END_IF;
                     END_IF;

                     #tempLengthIndex := #MODBUS_REQUEST_LENGTH;
                   END_REGION

                 #MB_FC_15_WRITE_COILS,
                 #MB_FC_16_WRITE_REGISTERS:
                   REGION 15 / 16 Write Coils / Registers
                     // write start address to array
                     #tempStartAddress := UINT_TO_WORD(#statStartAddress);
                     #statTransmitterBuffer[#MODBUS_STARTADDRESS_INDEX] := #tempStartAddress.%B1;
                     #statTransmitterBuffer[#MODBUS_STARTADDRESS_INDEX + #B1_OFFSET] := #tempStartAddress.%B0;

                     // write quantity to array
                     #tempQuantity := UINT_TO_WORD(#statQuantity);
                     #statTransmitterBuffer[#MODBUS_QUANTITY_INDEX] := #tempQuantity.%B1;
                     #statTransmitterBuffer[#MODBUS_QUANTITY_INDEX + #B1_OFFSET] := #tempQuantity.%B0;

                     // byte count 
                     #statTransmitterBuffer[#MODBUS_BYTE_COUNT_INDEX] := USINT_TO_BYTE(#statQuantityInBytes);

                     IF IS_ARRAY(#data) AND
                       (TypeOfElements(#data) = Byte OR TypeOfElements(#data) = Char)
                     THEN
                       // for an array at INOUT data MOVE_BLK_VARIANT is used to copy data from static receive buffer to the INOUT
                       #tempRetVal := MOVE_BLK_VARIANT(SRC := #data,
                                                       COUNT := #statQuantityInBytes,
                                                       SRC_INDEX := #DATA_INDEX_0,
                                                       DEST_INDEX := #MODBUS_DATA_INDEX,
                                                       DEST => #statTransmitterBuffer);
                       // if MOVE_BLK_VARIANT was executed with error, jump to AutoCleard error and give feedback to the user
                       IF #tempRetVal <> 0 THEN
                         #statErrorAutoCleared := TRUE;
                         #statDiagnostics.status := #ERR_MOVE_BLK_VAR_MULTIPLE_WRITE;
                         #statDiagnostics.subFunctionStatus := INT_TO_WORD(#tempRetVal);
                         #statDiagnostics.stateNumber := #statFBState;
                       END_IF;

                     ELSE
                       #tempSerializePos := #MODBUS_DATA_INDEX;
                       // for a structure or other datatype at INOUT data serialized is used to copy data from static receive buffer to the INOUT
                       #tempRetVal := Serialize(SRC_VARIABLE := #data,
                                                DEST_ARRAY => #statTransmitterBuffer,
                                                POS := #tempSerializePos);
                       // if serialize function was executed with error, jump to AutoCleared error and give feedback to the user
                       IF #tempRetVal <> 0 THEN
                         #statErrorAutoCleared := TRUE;
                         #statDiagnostics.status := #ERR_SERIALIZE_MULTIPLE_WRITE;
                         #statDiagnostics.subFunctionStatus := INT_TO_WORD(#tempRetVal);
                         #statDiagnostics.stateNumber := #statFBState;
                       END_IF;
                     END_IF;

                     #tempLengthIndex := #MODBUS_REQUEST_MULTIPLE_WRITE_LENGTH + #statQuantityInBytes;
                   END_REGION

                 #MB_FC_07_READ_EXCEPTION_STATUS:
                   REGION 07 Read Exception status
                     (*
                       This function code is used to read the contents of eight Exception Status outputs in a remote
                       device. Only address and function code needed
                     *)
                     #tempLengthIndex := #MODBUS_DEFAULT_REQUEST_LENGTH;
                   END_REGION 07 Read Exception status

                 #MB_FC_08_DIAGNOSTIC:
                   REGION 08 Diagnostics
                     // sub-function code (2Bytes) 2 X 2Bytes
                     // write sub-function code to to array
                     #tempStartAddress := UINT_TO_WORD(#statStartAddress);
                     #statTransmitterBuffer[#MODBUS_DIAG_SUB_FC_INDEX] := #tempStartAddress.%B1;
                     #statTransmitterBuffer[#MODBUS_DIAG_SUB_FC_INDEX + #B1_OFFSET] := #tempStartAddress.%B0;

                     CASE #statStartAddress OF
                       #DIAG_SUB_FC_0_RETURN_QUERY_DATA:
                         REGION Sub Function 00 - Return Query Data
                           // request sends two bytes, that have to be echoed by the slave
                           #tempQuantity := UINT_TO_WORD(#statQuantity);
                           #statTransmitterBuffer[#MODBUS_DIAG_DATA_INDEX] := #tempQuantity.%B1;
                           #statTransmitterBuffer[#MODBUS_DIAG_DATA_INDEX + #B1_OFFSET] := #tempQuantity.%B0;
                         END_REGION Sub Function 00 - Return Query #data

                       #DIAG_SUB_FC_1_RESTART_COM:
                         REGION Sub Function 01 - Restart Communication
                           // request data can be: 16#00 00 (leave log) or 16#FF 00 (clear log)
                           #tempQuantity := UINT_TO_WORD(#statQuantity);
                           IF #tempQuantity = 16#0000 OR #tempQuantity = #FC05_SET_COMMAND_IDENT THEN
                             #statTransmitterBuffer[#MODBUS_DIAG_DATA_INDEX] := #tempQuantity.%B1;
                             #statTransmitterBuffer[#MODBUS_DIAG_DATA_INDEX + #B1_OFFSET] := #tempQuantity.%B0;
                           ELSE
                             #statErrorAutoCleared := TRUE;
                             #statDiagnostics.status := #ERR_REQUEST_NOT_SUPPORTED_FUNCTION_CODE; // set correct status that identifies error clearly
                             #statDiagnostics.subFunctionStatus := USINT_TO_WORD(#statFunctionCode); // given function code
                             #statDiagnostics.stateNumber := #statFBState; // set error state number for diagnostic
                             EXIT; // leave state machine and its sourounding loop immediately
                           END_IF;
                         END_REGION Sub Function 01 - Restart Communication

                       #DIAG_SUB_FC_2_RETURN_DIAG_REGISTER,
                       #DIAG_SUB_FC_4_FORCE_LISTEN_ONLY,
                       #DIAG_SUB_FC_10_CLEAR_DIAG_REGISTER,
                       #DIAG_SUB_FC_11_COUNTER_TOTAL_MESSAGE,
                       #DIAG_SUB_FC_12_COUNTER_CRC_ERR,
                       #DIAG_SUB_FC_13_COUNTER_EXCEPTION_ERR,
                       #DIAG_SUB_FC_14_COUNTER_TOTAL_MESSAGES,
                       #DIAG_SUB_FC_15_COUNTER_NO_RESPONSE,
                       #DIAG_SUB_FC_16_COUNTER_NAK,
                       #DIAG_SUB_FC_17_COUNTER_SERVER_BUSY,
                       #DIAG_SUB_FC_18_BUS_CHAR_OVERRUN,
                       #DIAG_SUB_FC_20_CLEAR_OVERRUN:
                         (*
                           Request to get a counter of all information that the devices processed
                           since last restart or reset (sub-function code 10).
                           Sub-function code 4 request to acitivate listen only mode --> no responses will be given to Master.
                           The only function that is processed is FC 08 Sub-FC 01 to restart the communication of the slave.
                         *)
                         #statTransmitterBuffer[#MODBUS_DIAG_DATA_INDEX] := 16#00;
                         #statTransmitterBuffer[#MODBUS_DIAG_DATA_INDEX + #B1_OFFSET] := 16#00;

                       ELSE
                         // not supported Subfunction code for diagnostics is requested
                         #statErrorAutoCleared := TRUE;
                         #statDiagnostics.status := #ERR_NOT_SUPPORTED_SUB_FC;
                         #statDiagnostics.subFunctionStatus := UINT_TO_WORD(#statStartAddress);
                         #statDiagnostics.stateNumber := #statFBState;
                         EXIT;
                     END_CASE;
                     // set request length for ASCII encoding
                     #tempLengthIndex := #MODBUS_REQUEST_LENGTH;


                   END_REGION

                 #MB_FC_11_GET_COM_EVENT_COUNTER:
                   REGION 11 Get Communication Event Counter
                     (*
                       This function code is used to get a status word and an event count from the remote device's communication 
                       event counter.
                     *)
                     #tempLengthIndex := #MODBUS_DEFAULT_REQUEST_LENGTH;
                   END_REGION 11 Get Communication Event Counter

                 #MB_FC_12_GET_COM_EVENT_LOG:
                   REGION 12 Get Communication Event Log
                     (*
                       This function code is used to get a status word, event count, message count, and a field of
                       event bytes from the remote device.
                     *)
                     #tempLengthIndex := #MODBUS_DEFAULT_REQUEST_LENGTH;
                   END_REGION 12 Get Communication Event Log

                 #MB_FC_22_MASK_WRITE_REGISTER:
                   REGION Mask Write Register
                     (*
                       Request:
                       Function code     1 Byte    0x16
                       Reference Address 2 Bytes   0x0000 to 0xFFFF
                       And_Mask          2 Bytes   0x0000 to 0xFFFF
                       Or_Mask           2 Bytes   0x0000 to 0xFFFF
                     *)
                     #tempStartAddress := UINT_TO_WORD(#statStartAddress);
                     #statTransmitterBuffer[#MODBUS_STARTADDRESS_INDEX] := #tempStartAddress.%B1;
                     #statTransmitterBuffer[#MODBUS_STARTADDRESS_INDEX + #B1_OFFSET] := #tempStartAddress.%B0;

                     #statTransmitterBuffer[#MODBUS_AND_MASK_INDEX] := #statAndMask.%B1;
                     #statTransmitterBuffer[#MODBUS_AND_MASK_INDEX + #B1_OFFSET] := #statAndMask.%B0;

                     #statTransmitterBuffer[#MODBUS_OR_MASK_INDEX] := #statOrMask.%B1;
                     #statTransmitterBuffer[#MODBUS_OR_MASK_INDEX + #B1_OFFSET] := #statOrMask.%B0;

                     #tempLengthIndex := #MODBUS_REQUEST_MASK_WRITE_LENGTH;
                   END_REGION Mask Write Register

                 #MB_FC_23_READ_WRITE_MULTIPLE_REGISTERS:
                   REGION 23 Read/Write Multiple registers
                     (*
                       Request:
                       Function code           1 Byte      0x17 
                       Read Starting Address   2 Bytes     0x0000 to 0xFFFF 
                       Quantity to Read        2 Bytes     0x0001 to 0x007D 
                       Write Starting Address  2 Bytes     0x0000 to 0xFFFF 
                       Quantity to Write       2 Bytes     0x0001 to 0X0079 
                       Write Byte Count        1 Byte      2 x N* 
                       Write Registers Value   N*x 2 Bytes 
                     *)
                     // read Starting Address
                     #tempStartAddress := UINT_TO_WORD(#statReadWrite.startAddressRead - #MODBUS_STARTADDRESS_CORRECTION);
                     #statTransmitterBuffer[#MODBUS_STARTADDRESS_INDEX] := #tempStartAddress.%B1;
                     #statTransmitterBuffer[#MODBUS_STARTADDRESS_INDEX + #B1_OFFSET] := #tempStartAddress.%B0;

                     // quantity to Read
                     #tempQuantity := UINT_TO_WORD(#statReadWrite.quantityRead);
                     #statTransmitterBuffer[#MODBUS_QUANTITY_INDEX] := #tempQuantity.%B1;
                     #statTransmitterBuffer[#MODBUS_QUANTITY_INDEX + #B1_OFFSET] := #tempQuantity.%B0;

                     // write Starting Address
                     #tempStartAddress := UINT_TO_WORD(#statReadWrite.startAddressWrite - #MODBUS_STARTADDRESS_CORRECTION);
                     #statTransmitterBuffer[#MODBUS_STARTADDRESS_FC23_WRITE_INDEX] := #tempStartAddress.%B1;
                     #statTransmitterBuffer[#MODBUS_STARTADDRESS_FC23_WRITE_INDEX + #B1_OFFSET] := #tempStartAddress.%B0;

                     // quantity to Write 
                     #tempQuantity := UINT_TO_WORD(#statReadWrite.quantityWrite);
                     #statTransmitterBuffer[#MODBUS_QUANTITY_FC23_WRITE_INDEX] := #tempQuantity.%B1;
                     #statTransmitterBuffer[#MODBUS_QUANTITY_FC23_WRITE_INDEX + #B1_OFFSET] := #tempQuantity.%B0;

                     // write Byte Count
                     #statTransmitterBuffer[#MODBUS_BYTE_COUNT_FC23_INDEX] := UINT_TO_BYTE(#statQuantityInBytesWrite);

                     IF IS_ARRAY(#data) AND
                       (TypeOfElements(#data) = Byte OR TypeOfElements(#data) = Char)
                     THEN
                       // for an array at INOUT data MOVE_BLK_VARIANT is used to copy data from static receive buffer to the INOUT
                       #tempRetVal := MOVE_BLK_VARIANT(SRC := #data,
                                                       COUNT := #statQuantityInBytesWrite,
                                                       SRC_INDEX := #DATA_INDEX_0,
                                                       DEST_INDEX := #MODBUS_FC23_DATA_INDEX,
                                                       DEST => #statTransmitterBuffer);
                       // if MOVE_BLK_VARIANT was executed with error, jump to AutoCleard error and give feedback to the user
                       IF #tempRetVal <> 0 THEN
                         #statErrorAutoCleared := TRUE;
                         #statDiagnostics.status := #ERR_MOVE_BLK_VAR_MULTIPLE_WRITE;
                         #statDiagnostics.subFunctionStatus := INT_TO_WORD(#tempRetVal);
                         #statDiagnostics.stateNumber := #statFBState;
                       END_IF;

                     ELSE
                       #tempSerializePos := #MODBUS_FC23_DATA_INDEX;
                       // for a structure or other datatype at INOUT data serialized is used to copy data from static receive buffer to the INOUT
                       #tempRetVal := Serialize(SRC_VARIABLE := #data,
                                                DEST_ARRAY => #statTransmitterBuffer,
                                                POS := #tempSerializePos);
                       // if serialize function was executed with error, jump to AutoCleared error and give feedback to the user
                       IF #tempRetVal <> 0 THEN
                         #statErrorAutoCleared := TRUE;
                         #statDiagnostics.status := #ERR_SERIALIZE_MULTIPLE_WRITE;
                         #statDiagnostics.subFunctionStatus := INT_TO_WORD(#tempRetVal);
                         #statDiagnostics.stateNumber := #statFBState;
                       END_IF;
                     END_IF;

                     #tempLengthIndex := #MODBUS_REQUEST_READ_WRITE_LENGTH + #statQuantityInBytesWrite;
                   END_REGION 23 Read/Write Multiple registers

                 #MB_FC_43_READ_DEVICE_IDENT:
                   REGION 43 Read Device Identification
                     // FC 43 Read Device Identificaton
                     // MEI Type := 0E
                     // read Device ID code 01 (Basic) / 02 (regular) / 03 (extended) / 04 (specific)
                     // object ID (00 to FF)
                     // - 00 Vendor name (Mandatory) - BASIC
                     // - 01 Product code (Mandatory) - BASIC
                     // - 02 MajorMinorRevision (Mandatory) - BASIC
                     // - 03 Vendor URL (optional) - REGULAR
                     // - 04 ProductName (optional) - REGULAR
                     // - 05 ModelName (optional) - REGULAR
                     // - 06 UserApplicationName (optional) - REGULAR
                     // - 07-7F reserved (optional) - REGULAR
                     // - 80-FF (optional) - EXTENDED

                     // 16#08 for MEI Type Read Device Identification
                     #statTransmitterBuffer[#MODBUS_DIAG_SUB_FC_INDEX] := #MODBUS_FC43_MEI_TYE;
                     #tempStartAddress := UINT_TO_WORD(#statStartAddress);
                     // write to array
                     // read Device ID code 16#01 basic, 16#02 regular, 16#03 extended or 16#04 special identification object
                     #statTransmitterBuffer[#MODBUS_FC43_DEVICE_ID_CODE_INDEX] := #tempStartAddress.%B1;
                     // object ID 16#00 16#FF
                     #statTransmitterBuffer[#MODBUS_FC43_OBJECT_ID_CODE_INDEX] := #tempStartAddress.%B0;

                     #tempLengthIndex := #MODBUS_FC43_REQUEST_LENGTH;
                   END_REGION

                 ELSE // function code not supported
                   // write diagnostic Information
                   #statErrorAutoCleared := TRUE;
                   #statDiagnostics.status := #ERR_REQUEST_NOT_SUPPORTED_FUNCTION_CODE; // Set correct status that identifies error clearly
                   #statDiagnostics.subFunctionStatus := USINT_TO_WORD(#statFunctionCode); // Given function code
                   #statDiagnostics.stateNumber := #statFBState; // Set error state number for diagnostic
                   EXIT; // leave state machine and its sourounding loop immediately
               END_CASE;
             END_REGION Setup function code specific part

             // generate encoded ASCII protocol array
             #instAsciiEncode(lengthToConvert := #tempLengthIndex,
                              lengthConverted => #statLengthAfterEncoding,
                              binaryData := #statTransmitterBuffer,
                              asciiMessageData := #statTransmitterAsciiBuffer);

             // next state - start transmit
             #statFBState := #FB_STATE_TRANSMIT_DATA;
             // set repeat condition to TRUE to stay in lstatemaschine one more step
             #tempStayInStatemachine := TRUE;
           END_REGION Setup Transmit Protocol

         #FB_STATE_TRANSMIT_DATA:
           REGION Transmit data to slave
             // call transmission instance to transfer the request to the client / slave
             #instSendRequest(REQ := TRUE,
                              "PORT" := #statHardwareId,
                              LENGTH := DINT_TO_UINT(#statLengthAfterEncoding),
                              BUFFER := #statTransmitterAsciiBuffer);

             // transmission finished successfully
             IF (#instSendRequest.DONE = TRUE) THEN
               #instSendRequest(REQ := FALSE,
                                BUFFER := #statTransmitterAsciiBuffer);  // reset receiver config REQ input after call

               // set next state
               IF #statFunctionCode = #MB_FC_08_DIAGNOSTIC AND #statStartAddress = #DIAG_SUB_FC_4_FORCE_LISTEN_ONLY THEN
                 #statDone := TRUE;
                 #statBusy := FALSE;
                 #statTransmitterBuffer := #tempEmptyData;
                 FILL_BLK(IN:=16#00,
                          COUNT:=DINT_TO_UINT(#BUFFER_UPPER_BOUND_ASCII + 1),
                          OUT=>#statTransmitterAsciiBuffer[0]);
                 #statDiagnostics.status := #STATUS_DONE;
                 #statFBState := #FB_STATE_WAIT_FOR_EXECUTE;
               ELSE
                 IF #statSlaveAddress = #MODBUS_ADDRESS_BROADCAST THEN
                   // if broadcast was send, go to delay turnaround
                   #statFBState := #FB_STATE_WAIT_FOR_TURNAROUND_DELAY;
                 ELSE
                   // if regular client was called, go to "wait for response"
                   #statFBState := #FB_STATE_WAIT_FOR_RESPONSE;
                 END_IF;
               END_IF;

               // reset watchdog previously to monitor time out of reception / tournaround delay
               #instWatchdog.TON(IN := FALSE,
                                 PT := #statParameter.transmissionWatchdog);

               // error occurred during data transmission
             ELSIF (#instSendRequest.ERROR = TRUE) THEN
               // write diagnostic Information
               #statErrorAutoCleared := TRUE;
               #statDiagnostics.status := #ERR_TRANSMISSION_FAILURE; // Set correct status that identifies error clearly
               #statDiagnostics.subFunctionStatus := #instSendRequest.STATUS; // Status of transmission instance
               #statDiagnostics.stateNumber := #statFBState; // Set error state number for diagnostic

               #instSendRequest(REQ := FALSE,
                                BUFFER := #statTransmitterAsciiBuffer);
             END_IF;
           END_REGION Transmit data to slave

         #FB_STATE_WAIT_FOR_TURNAROUND_DELAY:
           REGION Wait for TurnAround delay after Broadcast message
             // start watchdog to monitor time out of reception
             #instWatchdog.TON(IN := TRUE,
                               PT := #MODBUS_TURNAROUND_DELAY);

             // after reaching the TournAround time, exit block for next call
             IF #instWatchdog.Q = TRUE THEN
               #statDiagnostics.status := #STATUS_DONE;
               #statDone := TRUE;
               #statBusy := FALSE;
               #statFBState := #FB_STATE_WAIT_FOR_EXECUTE;
             END_IF;
           END_REGION Wait for TurnAround delay after Broadcast message

         #FB_STATE_WAIT_FOR_RESPONSE:
           REGION Wait for response from slave
             // call receiver instance to wait for incoming respose data
             #instGetResponse("PORT" := #statHardwareId,
                           BUFFER := #statReceiverAsciiBuffer);

             // start watchdog to monitor time out of reception
             #instWatchdog.TON(IN := TRUE,
                               PT := #statParameter.transmissionWatchdog);

             // port configuration finished successfully
             IF (#instGetResponse.NDR = TRUE) THEN
               // decode from ASCII to Byte Array
               #instAsciiDecode(lengthToDecode := #instGetResponse.LENGTH,
                                lengthConverted => #statLengthAfterDecoding,
                                asciiMessageData := #statReceiverAsciiBuffer,
                                binaryData := #statReceiverBuffer);

               IF #instAsciiDecode.resultOfLrcCheck = TRUE AND #instAsciiDecode.error = FALSE THEN
                 // set next state
                 #statFBState := #FB_STATE_PROCESS_RECEIVED_DATA;
                 #tempStayInStatemachine := TRUE;
               ELSE
                 // if error happend but retry counter greater than zero
                 IF (#statRetryCounter > 0) THEN
                   // decrement retry counter
                   #statRetryCounter -= 1;
                   // go back to transmittion and start a retransmittion
                   #statFBState := #FB_STATE_TRANSMIT_DATA;
                 ELSE
                   // write diagnostic Information
                   #statErrorAutoCleared := TRUE;
                   #statDiagnostics.subFunctionStatus := #NO_ERROR; // no subfunction status
                   #statDiagnostics.stateNumber := #statFBState; // set error state number for diagnostic
                   IF #instAsciiDecode.resultOfLrcCheck = FALSE AND #instAsciiDecode.error = FALSE THEN
                     #statDiagnostics.status := #ERR_RESPONSE_WRONG_LRC; // set correct status that identifies error clearly
                   ELSE
                     #statDiagnostics.status := #ERR_TRANSMISSION_FAILURE; // set correct status that identifies error clearly
                   END_IF;
                 END_IF;
               END_IF;

               // error occurred during data reception
             ELSIF (#instGetResponse.ERROR = TRUE) THEN
               // check if retry counter is greater than zeror --> retry transmission
               IF (#statRetryCounter > 0) THEN
                 // decrement retry counter
                 #statRetryCounter -= 1;
                 // go back to transmittion and start a retransmittion
                 #statFBState := #FB_STATE_TRANSMIT_DATA;
               ELSE
                 // write diagnostic Information
                 #statErrorAutoCleared := TRUE;
                 #statDiagnostics.status := #ERR_RECEIVER_FAILURE; // set correct status that identifies error clearly
                 #statDiagnostics.subFunctionStatus := #instGetResponse.STATUS; // status of Port Configuration
                 #statDiagnostics.stateNumber := #statFBState; // set error state number for diagnostic
               END_IF;

               // if watchdog time is expired / reached its time, return error and end Block call
             ELSIF (#instWatchdog.Q = TRUE) THEN
               // check id retry counter is greater than zeror --> retry transmission
               IF (#statRetryCounter > 0) THEN
                 // decrement retry counter
                 #statRetryCounter -= 1;
                 // go back to transmittion and start a retransmittion
                 #statFBState := #FB_STATE_TRANSMIT_DATA;
               ELSE
                 // write diagnostic Information
                 #statErrorAutoCleared := TRUE;
                 #statDiagnostics.status := #ERR_RESPONSE_TIMEOUT_EXPIRATION; // set correct status that identifies error clearly
                 #statDiagnostics.subFunctionStatus := #NO_ERROR; // no subfunction status
                 #statDiagnostics.stateNumber := #statFBState; // set error state number for diagnostic
               END_IF;
             END_IF;
           END_REGION Wait for response from slave

         #FB_STATE_PROCESS_RECEIVED_DATA: // further processing state
           REGION Process received data
             IF #statReceiverBuffer[#MODBUS_SLAVE_ADDRESS_INDEX] <> USINT_TO_BYTE(#statSlaveAddress) THEN
               // write diagnostic Information
               #statErrorAutoCleared := TRUE;
               #statDiagnostics.status := #ERR_RESPONSE_WRONG_SLAVE; // set correct status that identifies error clearly
               #statDiagnostics.subFunctionStatus := #statReceiverBuffer[#MODBUS_SLAVE_ADDRESS_INDEX]; // slave address of response that was received
               #statDiagnostics.stateNumber := #statFBState; // set error state number for diagnostic

               // check response for error / exeption --> MSB of FunctionCode 0x8...
             ELSIF #statReceiverBuffer[#MODBUS_EXCEPTION_CODE_INDEX].%X7 = TRUE THEN
               // write diagnostic Information
               #statErrorAutoCleared := TRUE;
               #statDiagnostics.status := #ERR_RESPONSE_EXCEPTION_FROM_SLAVE; // set correct status that identifies error clearly
               #statDiagnostics.subFunctionStatus.%B1 := #statReceiverBuffer[#MODBUS_EXCEPTION_CODE_INDEX]; // exception code of Modbus protocol
               #statDiagnostics.subFunctionStatus.%B0 := #statReceiverBuffer[#MODBUS_EXCEPTION_CODE_INDEX + #B1_OFFSET]; // error info of Modbus protocol
               #statDiagnostics.stateNumber := #statFBState; // set error state number for diagnostic

             ELSE

               REGION Decode functioncode specific response
                 // every responses first byte is the function code, check if it matches to the requested FC
                 IF BYTE_TO_USINT(#statReceiverBuffer[#MODBUS_FUNCTION_CODE_INDEX]) <> #statFunctionCode THEN
                   // requested function code does not match to the requested
                   #statErrorAutoCleared := TRUE;
                   #statDiagnostics.status := #ERR_RESPONSE_NOT_EXPECTED_FC; // Set correct status that identifies error clearly
                   #statDiagnostics.subFunctionStatus := USINT_TO_WORD(#statFunctionCode);
                   #statDiagnostics.stateNumber := #statFBState; // Set error state number for diagnostic
                   EXIT; // leave state machine and its sourounding loop immediately
                 ELSE
                   // correct FC had been received, further information can be decoded
                   CASE #statFunctionCode OF
                     #MB_FC_01_READ_COILS,
                     #MB_FC_02_READ_DISCRETE_INPUTS,
                     #MB_FC_03_READ_HOLDING_REGISTERS,
                     #MB_FC_04_READ_INPUT_REGISTERS:
                       REGION 01 / 02 / 03 / 04 check length
                         // response contains function code and Byte count
                         // check if byte count  and function code match with the request
                         IF BYTE_TO_USINT(#statReceiverBuffer[#MODBUS_RESPONSE_BYTE_COUNT_INDEX]) > #statQuantityInBytes THEN
                           // requested length does not match to the length, that was received
                           #statErrorAutoCleared := TRUE;
                           #statDiagnostics.status := #ERR_RESPONSE_WRONG_QUANTITY; // set correct status that identifies error clearly
                           #statDiagnostics.subFunctionStatus := USINT_TO_WORD(#statFunctionCode);
                           #statDiagnostics.stateNumber := #statFBState; // set error state number for diagnostic
                           EXIT; // leave state machine and its sourounding loop immediately
                         END_IF;
                         #tempReceiveBufferIndex := #MODBUS_USER_DATA_READ_INDEX;

                       END_REGION

                     #MB_FC_05_WRITE_COIL,
                     #MB_FC_06_WRITE_REGISTER:
                       REGION 05 / 06 check response of writing single coil / register
                         // response code contains functon code, output address and output value
                         //check if the request matches with the response
                         #tempStartAddress := UINT_TO_WORD(#statStartAddress);
                         IF #statReceiverBuffer[#MODBUS_RESPONSE_ADDRESS_INDEX] <> #tempStartAddress.%B1
                           OR #statReceiverBuffer[#MODBUS_RESPONSE_ADDRESS_INDEX + #B1_OFFSET] <> #tempStartAddress.%B0
                           OR #statReceiverBuffer[#MODBUS_RESPONSE_QUANTITY_INDEX] <> #statTransmitterBuffer[#MODBUS_QUANTITY_INDEX]
                           OR #statReceiverBuffer[#MODBUS_RESPONSE_QUANTITY_INDEX + #B1_OFFSET] <> #statTransmitterBuffer[#MODBUS_QUANTITY_INDEX + #B1_OFFSET]
                         THEN
                           #statErrorAutoCleared := TRUE;
                           #statDiagnostics.status := #ERR_RESPONSE_SINGLE_WRITE; // Set correct status that identifies error clearly
                           #statDiagnostics.subFunctionStatus := USINT_TO_WORD(#statFunctionCode);
                           #statDiagnostics.stateNumber := #statFBState; // Set error state number for diagnostic
                           EXIT; // leave state machine and its sourounding loop immediately
                         END_IF;

                       END_REGION

                     #MB_FC_15_WRITE_COILS,
                     #MB_FC_16_WRITE_REGISTERS:
                       REGION 15 / 16 check response of wrting Write Coils and registers
                         // response code contains function code, output address and quantity of outputs
                         // check if the request matches with the response
                         #tempStartAddress := UINT_TO_WORD(#statStartAddress);
                         IF #statReceiverBuffer[#MODBUS_RESPONSE_ADDRESS_INDEX] <> #tempStartAddress.%B1
                             OR #statReceiverBuffer[#MODBUS_RESPONSE_ADDRESS_INDEX + #B1_OFFSET] <> #tempStartAddress.%B0
                             OR #statReceiverBuffer[#MODBUS_RESPONSE_QUANTITY_INDEX] <> #statTransmitterBuffer[#MODBUS_QUANTITY_INDEX]
                             OR #statReceiverBuffer[#MODBUS_RESPONSE_QUANTITY_INDEX + #B1_OFFSET] <> #statTransmitterBuffer[#MODBUS_QUANTITY_INDEX + #B1_OFFSET]
                         THEN
                           #statErrorAutoCleared := TRUE;
                           #statDiagnostics.status := #ERR_RESPONSE_MULTI_WRITE; // set correct status that identifies error clearly
                           #statDiagnostics.subFunctionStatus := USINT_TO_WORD(#statFunctionCode);
                           #statDiagnostics.stateNumber := #statFBState; // set error state number for diagnostic
                           EXIT; // leave state machine and its sourounding loop immediately
                         END_IF;
                       END_REGION

                     #MB_FC_07_READ_EXCEPTION_STATUS:
                       REGION Read Exception Status
                         #tempReceiveBufferIndex := #MODBUS_DEFAULT_RESP_INDEX;
                       END_REGION Read Exception Status

                     #MB_FC_08_DIAGNOSTIC:
                       REGION 08 Diagnostics
                         // response code contains function code, subfunction code and subfunction data (depending on subfunction)
                         // check which subfunction was requested and check data
                         // check if the request matches with the response
                         #tempStartAddress := UINT_TO_WORD(#statStartAddress);
                         IF #statReceiverBuffer[#MODBUS_DIAG_SUB_FC_INDEX] <> #tempStartAddress.%B1
                           OR #statReceiverBuffer[#MODBUS_DIAG_SUB_FC_INDEX + #B1_OFFSET] <> #tempStartAddress.%B0
                         THEN
                           #statErrorAutoCleared := TRUE;
                           #statDiagnostics.status := #ERR_RESPONSE_NOT_EXPECTED_SUB_FC; // set correct status that identifies error clearly
                           #statDiagnostics.subFunctionStatus := USINT_TO_WORD(#statFunctionCode);
                           #statDiagnostics.stateNumber := #statFBState; // set error state number for diagnostic
                           EXIT; // leave state machine and its sourounding loop immediately
                         END_IF;

                         CASE WORD_TO_USINT(#tempStartAddress) OF
                           #DIAG_SUB_FC_0_RETURN_QUERY_DATA:
                             REGION Sub Function 00 - Return Query Data
                               #tempQuantity.%B1 := #statReceiverBuffer[#MODBUS_DIAG_DATA_INDEX];
                               #tempQuantity.%B0 := #statReceiverBuffer[#MODBUS_DIAG_DATA_INDEX + #B1_OFFSET];
                               IF WORD_TO_UINT(#tempQuantity) <> #statQuantity THEN
                                 #statErrorAutoCleared := TRUE;
                                 #statDiagnostics.status := #ERR_DIAG_SUB_0; // set correct status that identifies error clearly
                                 #statDiagnostics.subFunctionStatus := #tempQuantity;  // wrong Echo value
                                 #statDiagnostics.stateNumber := #statFBState; // set error state number for diagnostic
                                 EXIT; // leave state machine and its sourounding loop immediately
                               ELSE
                                 #tempReceiveBufferIndex := #MODBUS_DIAG_DATA_INDEX;
                               END_IF;
                             END_REGION Sub Function 00 - Return Query Data

                           #DIAG_SUB_FC_1_RESTART_COM:
                             REGION Sub Function 01 - Restart Communication
                               // response contains echo of request data 00 (leave log) / FF (clear log)
                               #tempQuantity.%B1 := #statReceiverBuffer[#MODBUS_DIAG_DATA_INDEX];
                               #tempQuantity.%B0 := #statReceiverBuffer[#MODBUS_DIAG_DATA_INDEX + #B1_OFFSET];
                               IF WORD_TO_UINT(#tempQuantity) <> #statQuantity THEN
                                 #statErrorAutoCleared := TRUE;
                                 #statDiagnostics.status := #ERR_DIAG_SUB_1; // set correct status that identifies error clearly
                                 #statDiagnostics.subFunctionStatus := #tempQuantity;  // wrong Echo value
                                 #statDiagnostics.stateNumber := #statFBState; // set error state number for diagnostic
                                 EXIT; // leave state machine and its sourounding loop immediately
                               ELSE
                                 #tempReceiveBufferIndex := #MODBUS_DIAG_DATA_INDEX;
                               END_IF;
                             END_REGION Sub Function 01 - Restart Communication

                           #DIAG_SUB_FC_10_CLEAR_DIAG_REGISTER:
                             REGION Sub Function 10 - Clear Diag Register
                               // response contains echo of request data
                               IF #statReceiverBuffer[#MODBUS_DIAG_DATA_INDEX] <> #statTransmitterBuffer[#MODBUS_DIAG_DATA_INDEX]
                                 OR #statReceiverBuffer[#MODBUS_DIAG_DATA_INDEX + #B1_OFFSET] <> #statTransmitterBuffer[#MODBUS_DIAG_DATA_INDEX + #B1_OFFSET]
                               THEN
                                 #statErrorAutoCleared := TRUE;
                                 #statDiagnostics.status := #ERR_DIAG_SUB_0; // set correct status that identifies error clearly
                                 #statDiagnostics.subFunctionStatus.%B1 := #statReceiverBuffer[#MODBUS_DIAG_DATA_INDEX];
                                 #statDiagnostics.subFunctionStatus.%B0 := #statReceiverBuffer[#MODBUS_DIAG_DATA_INDEX + #B1_OFFSET];
                                 #statDiagnostics.stateNumber := #statFBState; // set error state number for diagnostic
                                 EXIT; // leave state machine and its sourounding loop immediately
                               ELSE
                                 #tempReceiveBufferIndex := #MODBUS_DIAG_DATA_INDEX;
                               END_IF;
                             END_REGION Sub Function 10 - Clear Diag Register

                           #DIAG_SUB_FC_4_FORCE_LISTEN_ONLY:
                             // no response returned --> listen only mode (can only be restarted by FC 08 SUB FC 01)
                             ;

                           #DIAG_SUB_FC_2_RETURN_DIAG_REGISTER,
                           // response contains diagnostic register contents 
                           #DIAG_SUB_FC_11_COUNTER_TOTAL_MESSAGE,
                           // response contains total message count of modbus slave
                           #DIAG_SUB_FC_12_COUNTER_CRC_ERR,
                           // response contains CRC error count of modbus slave
                           #DIAG_SUB_FC_13_COUNTER_EXCEPTION_ERR,
                           // response contains exception error count of modbus slave
                           #DIAG_SUB_FC_14_COUNTER_TOTAL_MESSAGES,
                           // response contains server message count of modbus slave
                           #DIAG_SUB_FC_15_COUNTER_NO_RESPONSE,
                           // response contains server no response count of modbus slave
                           #DIAG_SUB_FC_16_COUNTER_NAK,
                           // response contains server Negative Acknowledge (NAK)count of modbus slave
                           #DIAG_SUB_FC_17_COUNTER_SERVER_BUSY:
                             // response contains server device busy count of modbus slave
                             // always same data length, which content can not be known before, so just copying to INOUT data
                             #tempReceiveBufferIndex := #MODBUS_DIAG_DATA_INDEX;
                           ELSE  // statement section ELSE
                             ;
                         END_CASE;

                       END_REGION

                     #MB_FC_11_GET_COM_EVENT_COUNTER:
                       REGION Get Comm Event Counter
                         #tempReceiveBufferIndex := #MODBUS_DEFAULT_RESP_INDEX;
                       END_REGION Get Comm Event Counter

                     #MB_FC_12_GET_COM_EVENT_LOG:
                       REGION Get Comm Event Log
                         #tempReceiveBufferIndex := #MODBUS_DEFAULT_RESP_INDEX + 1;
                         #statQuantityInBytes := BYTE_TO_USINT(#statReceiverBuffer[#MODBUS_DEFAULT_RESP_INDEX]);
                       END_REGION Get Comm Event Log

                     #MB_FC_22_MASK_WRITE_REGISTER:
                       REGION 22 Mask Write Register - check response of mask request
                         // response code contains functon code, output address and output value
                         // check if the request matches with the response
                         #tempStartAddress := UINT_TO_WORD(#statStartAddress);
                         IF #statReceiverBuffer[#MODBUS_STARTADDRESS_INDEX] <> #tempStartAddress.%B1
                           OR #statReceiverBuffer[#MODBUS_STARTADDRESS_INDEX + #B1_OFFSET] <> #tempStartAddress.%B0
                           OR #statReceiverBuffer[#MODBUS_AND_MASK_INDEX] <> #statTransmitterBuffer[#MODBUS_AND_MASK_INDEX]
                           OR #statReceiverBuffer[#MODBUS_AND_MASK_INDEX + #B1_OFFSET] <> #statTransmitterBuffer[#MODBUS_AND_MASK_INDEX + #B1_OFFSET]
                           OR #statReceiverBuffer[#MODBUS_OR_MASK_INDEX] <> #statTransmitterBuffer[#MODBUS_OR_MASK_INDEX]
                           OR #statReceiverBuffer[#MODBUS_OR_MASK_INDEX + #B1_OFFSET] <> #statTransmitterBuffer[#MODBUS_OR_MASK_INDEX + #B1_OFFSET]
                         THEN
                           #statErrorAutoCleared := TRUE;
                           #statDiagnostics.status := #ERR_RESPONSE_SINGLE_WRITE; // set correct status that identifies error clearly
                           #statDiagnostics.subFunctionStatus := USINT_TO_WORD(#statFunctionCode);
                           #statDiagnostics.stateNumber := #statFBState; // set error state number for diagnostic
                           EXIT; // leave state machine and its sourounding loop immediately
                         END_IF;
                       END_REGION 22 Mask Write Register - check response of mask request

                     #MB_FC_23_READ_WRITE_MULTIPLE_REGISTERS:
                       REGION 23 Read/Write Multiple registers - check length
                         // response contains function code and Byte count
                         // check if byte count  and function code match with the request
                         IF BYTE_TO_USINT(#statReceiverBuffer[#MODBUS_FUNCTION_CODE_INDEX + #B1_OFFSET]) > #statQuantityInBytesRead THEN
                           // requested length does not match to the length, that was received
                           #statErrorAutoCleared := TRUE;
                           #statDiagnostics.status := #ERR_RESPONSE_WRONG_QUANTITY; // set correct status that identifies error clearly
                           #statDiagnostics.subFunctionStatus := USINT_TO_WORD(#statFunctionCode);
                           #statDiagnostics.stateNumber := #statFBState; // set error state number for diagnostic
                           EXIT; // leave state machine and its sourounding loop immediately
                         ELSE
                           #statQuantityInBytes := #statQuantityInBytesRead;
                         END_IF;
                         #tempReceiveBufferIndex := #MODBUS_USER_DATA_READ_INDEX;

                       END_REGION

                     #MB_FC_43_READ_DEVICE_IDENT:
                       REGION 43 Read Device Identification
                         // evaluation has to be done by user. Response is directly handed over to INOUT 'data'.
                         #tempReceiveBufferIndex := #MODBUS_DIAG_SUB_FC_INDEX;
                       END_REGION

                     ELSE // function code not supported
                       // write diagnostic Information
                       #statErrorAutoCleared := TRUE;
                       #statDiagnostics.status := #ERR_RESPONSE_NOT_SUPPORTED_FUNCTION_CODE; // set correct status that identifies error clearly
                       #statDiagnostics.subFunctionStatus := BYTE_TO_WORD(#statReceiverBuffer[#MODBUS_FUNCTION_CODE_INDEX]); // returned Function code
                       #statDiagnostics.stateNumber := #statFBState; // set error state number for diagnostic
                       EXIT; // leave state machine and its sourounding loop immediately
                   END_CASE;
                 END_IF;
               END_REGION Setup function code specific part

               // MOVE_BLK_VAR / Deserialize
               REGION Move received data
                 // data is just contained in the following Modbus function codes All others are done.
                 IF #statFunctionCode = #MB_FC_01_READ_COILS
                   OR #statFunctionCode = #MB_FC_02_READ_DISCRETE_INPUTS
                   OR #statFunctionCode = #MB_FC_03_READ_HOLDING_REGISTERS
                   OR #statFunctionCode = #MB_FC_04_READ_INPUT_REGISTERS
                   OR #statFunctionCode = #MB_FC_07_READ_EXCEPTION_STATUS
                   OR (#statFunctionCode = #MB_FC_08_DIAGNOSTIC AND #statQuantity <> #DIAG_SUB_FC_4_FORCE_LISTEN_ONLY)
                   OR #statFunctionCode = #MB_FC_12_GET_COM_EVENT_LOG
                   OR #statFunctionCode = #MB_FC_11_GET_COM_EVENT_COUNTER
                   OR #statFunctionCode = #MB_FC_23_READ_WRITE_MULTIPLE_REGISTERS
                   OR #statFunctionCode = #MB_FC_43_READ_DEVICE_IDENT
                 THEN
                   IF
                     IS_ARRAY(#data)
                     AND (TypeOfElements(#data) = Byte
                     OR TypeOfElements(#data) = Char)
                   THEN
                     // MOVE_VAR
                     #tempRetVal := MOVE_BLK_VARIANT(SRC := #statReceiverBuffer,
                                                     COUNT := #statQuantityInBytes,
                                                     SRC_INDEX := #tempReceiveBufferIndex,
                                                     DEST_INDEX := 0, DEST => #data);
                     // if MOVE_BLK_VARIANT was executed with error, jump to AutoCleared error and give feedback to the user
                     IF #tempRetVal <> 0 THEN
                       #statErrorAutoCleared := TRUE;
                       #statDiagnostics.status := #ERR_MOVE_BLK_VAR_RECEIVE_DATA;
                       #statDiagnostics.subFunctionStatus := INT_TO_WORD(#tempRetVal);
                       #statDiagnostics.stateNumber := #statFBState;
                     END_IF;
                   ELSE
                     #tempDeserializePos := #tempReceiveBufferIndex;
                     // for a structure or other datatype at INOUT data derserialized is used to copy data from static receive buffer to the INOUT
                     #tempRetVal := Deserialize(SRC_ARRAY := #statReceiverBuffer,
                                                DEST_VARIABLE => #data,
                                                POS := #tempDeserializePos);
                     // if Deserialize function was executed with error, jump to AutoCleared error and give feedback to the user
                     IF #tempRetVal <> 0 THEN
                       #statErrorAutoCleared := TRUE;
                       #statDiagnostics.status := #ERR_DESERIALIZE_TO_DATA;
                       #statDiagnostics.subFunctionStatus := INT_TO_WORD(#tempRetVal);
                       #statDiagnostics.stateNumber := #statFBState;
                     END_IF;
                   END_IF;

                 ELSE
                   // no data has to be copied for write, data is used for request data
                   ;
                 END_IF;

                 // end of Block
                 IF #tempRetVal = WORD_TO_INT(#NO_ERROR) THEN
                   #statDone := TRUE;
                   #statBusy := FALSE;
                   #statDiagnostics.status := #STATUS_DONE;
                   #statFBState := #FB_STATE_WAIT_FOR_EXECUTE;

                   REGION Clear Buffers
                     #statTransmitterBuffer := #tempEmptyData;
                     #statReceiverBuffer := #tempEmptyData;
                     FILL_BLK(IN := 16#00,
                              COUNT := DINT_TO_UINT(#BUFFER_UPPER_BOUND_ASCII + 1),
                              OUT => #statTransmitterAsciiBuffer[0]);
                     FILL_BLK(IN := 16#00,
                              COUNT := DINT_TO_UINT(#BUFFER_UPPER_BOUND_ASCII + 1),
                              OUT => #statReceiverAsciiBuffer[0]);
                   END_REGION Clear Buffers

                 END_IF;
               END_REGION ;
             END_IF;
           END_REGION Read and decode received data

         #FB_STATE_DISABLING:
           REGION Disabling
             // initialize all instances, if FB is disabled during any active instance.
             #instWatchdog.TON(IN := TRUE,
                               PT := #FB_DISABLE_TIME);
             #instSendRequest(REQ := FALSE,
                              BUFFER := #statTransmitterAsciiBuffer);
             #instPortConfig(REQ:=FALSE);
             #instTransmitterConfig(REQ := FALSE);
             #instReceiverConfig(REQ := FALSE,
                                 Receive_Conditions:=#statReceiverConditions);
             #instResetRxBuffer(REQ:=FALSE);

             IF (#instSendRequest.STATUS = #STATUS_NO_CALL AND
               #instPortConfig.STATUS = #STATUS_NO_CALL AND
               #instTransmitterConfig.STATUS = #STATUS_NO_CALL AND
               #instReceiverConfig.STATUS = #STATUS_NO_CALL AND
               #instResetRxBuffer.STATUS = #STATUS_NO_CALL)
               OR
               #instWatchdog.Q = TRUE
             THEN
               #statDisablingCompleted := TRUE;
               #statHardwareId := 0;
               #statFunctionCode := 0;
               #statSlaveAddress := 0;
               #statQuantity := 0;
               #statStartAddress := 0;
               #statAndMask := 0;
               #statOrMask := 0;

               // empty Data
               VariantPut(SRC := #tempEmptyData,
                          DST := #data);
             END_IF;
           END_REGION

         ELSE // undefined state in state machine reached
           #statDiagnostics.status := #ERR_UNDEFINED_STATE;
           #statDiagnostics.subFunctionStatus := #NO_ERROR;
           #statDiagnostics.stateNumber := #statFBState;
       END_CASE;
       // leave state machine or repeat if tag is set to TRUE by the user
     UNTIL #tempStayInStatemachine = FALSE END_REPEAT;
   END_REGION STATE_MACHINE

   REGION OUTPUTS
     // write outputs
     IF (#statDisablingCompleted = TRUE) THEN
       REGION disabling
         // reset outputs if disabling completed
         #statValid := FALSE;
         #statBusy := FALSE;
         #statError := FALSE;
         #statErrorUserCleared := FALSE;
         #statErrorAutoCleared := FALSE;
         #statDiagnostics.status := #STATUS_NO_CALL;
         #statDiagnostics.subFunctionStatus := #STATUS_DONE;
         #statDiagnostics.stateNumber := #FB_STATE_NO_PROCESSING_IDLE;
         #diagnostics := #statDiagnostics;
       END_REGION disabling

     ELSIF (#statErrorUserCleared = TRUE) AND (#statError = FALSE) THEN
       REGION error user cleared
         // error can only be cleared by user; rising edge at enable input is needed to continue 
         #statValid := FALSE;
         #statBusy := FALSE;
         #statError := TRUE;
         // write diagnostics
         #diagnostics.status := #statDiagnostics.status;
         #diagnostics.subFunctionStatus := #statDiagnostics.subFunctionStatus;
         #diagnostics.stateNumber := #statDiagnostics.stateNumber;
         #statFBState := #FB_STATE_NO_PROCESSING_IDLE;
       END_REGION error user cleared

     ELSIF (#statErrorAutoCleared = TRUE) AND (#statError = FALSE) THEN
       REGION error auto cleared
         // error can be reset by FB automatically
         #statDone := FALSE;
         #statValid := FALSE;
         #statBusy := FALSE;
         #statError := TRUE;
         // write diagnostics
         #diagnostics.status := #statDiagnostics.status;
         #diagnostics.subFunctionStatus := #statDiagnostics.subFunctionStatus;
         #diagnostics.stateNumber := #statDiagnostics.stateNumber;
         // go to wait for new execute
         #statErrorAutoCleared := FALSE;
         #statFBState := #FB_STATE_WAIT_FOR_EXECUTE;
       END_REGION error auto cleared

